(* IEC 61131-3 sources: plc-vscode/tests/st/all/rusty/tests/lit/multi/extern_C_fb_init, 1 file *)

(* ---- main.st ---- *)
FUNCTION main
VAR
    f: myFunctionBlock;
END_VAR
    printf('%d$N', f.a);
    printf('%d$N', f.b);
END_FUNCTION
